ORGANIZATION_BLOCK "Main"
VERSION : 0.1
BEGIN
	"FC_Used"();
END_ORGANIZATION_BLOCK

FUNCTION "FC_Used" : Void
VERSION : 0.1
BEGIN
	;
END_FUNCTION

FUNCTION "FC_Unused" : Void // PLCA-Q008
VERSION : 0.1
BEGIN
	;
END_FUNCTION
